{attribute 'qualified_only'}
{attribute 'strict'}
TYPE E_Ingredient_type :
(
	eNone := 0,
	eWater,
	ePowder,
	eOil
);
END_TYPE

(* stored: Version 1.1.0.1, ProductVersion 3.1.4024.15
   DUT E_Ingredient_type: Id {db9776dc-aa5e-4589-b841-68606adbf679} *)
